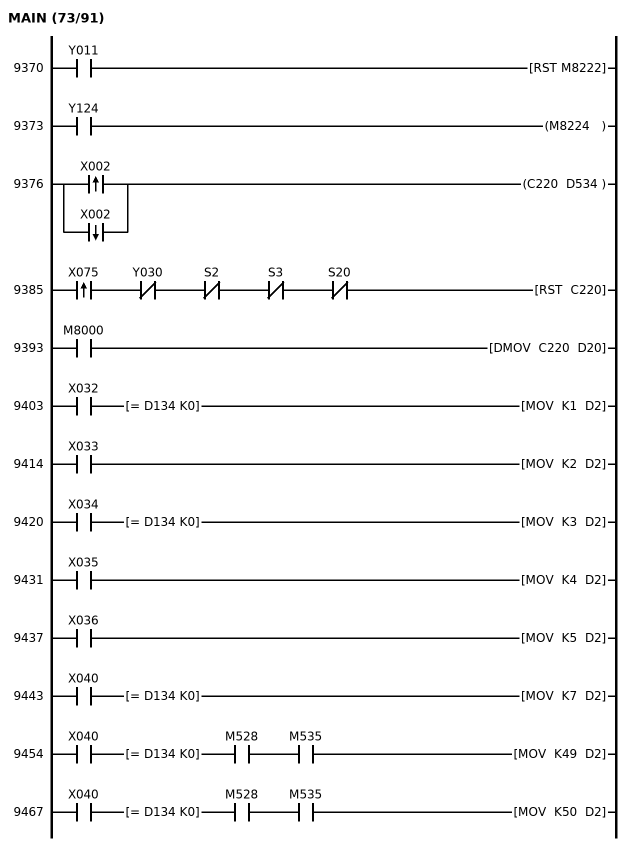
[picture p72: ladder of MAIN, rungs at steps 9370 to 9467]
9370  LD      Y011
      RST     M8222
9373  LD      Y124
      OUT     M8224
9376  LDP     X002
      ORF     X002
      OUT     C220 D534
9385  LDP     X075
      ANI     Y030
      ANI     S2
      ANI     S3
      ANI     S20
      RST     C220
9393  LD      M8000
      DMOV    C220 D20
9403  LD      X032
      AND=    D134 K0
      MOV     K1 D2
9414  LD      X033
      MOV     K2 D2
9420  LD      X034
      AND=    D134 K0
      MOV     K3 D2
9431  LD      X035
      MOV     K4 D2
9437  LD      X036
      MOV     K5 D2
9443  LD      X040
      AND=    D134 K0
      MOV     K7 D2
9454  LD      X040
      AND=    D134 K0
      AND     M528
      AND     M535
      MOV     K49 D2
9467  LD      X040
      AND=    D134 K0
      AND     M528
      AND     M535
      MOV     K50 D2
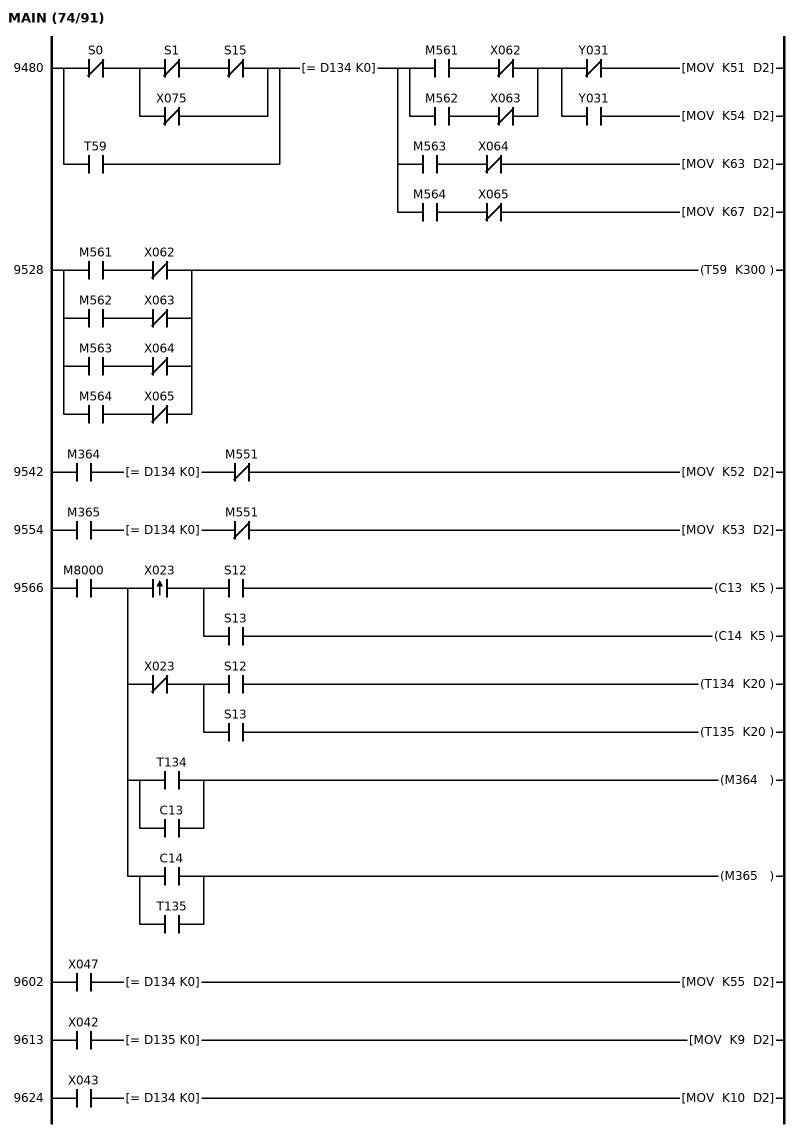
9480  LDI     S0
      LDI     S1
      ANI     S15
      ORI     X075
      ANB
      OR      T59
      AND=    D134 K0
      MPS
      LD      M561
      ANI     X062
      LD      M562
      ANI     X063
      ORB
      ANB
      MPS
      ANI     Y031
      MOV     K51 D2
      MPP
      AND     Y031
      MOV     K54 D2
      MRD
      AND     M563
      ANI     X064
      MOV     K63 D2
      MPP
      AND     M564
      ANI     X065
      MOV     K67 D2
9528  LD      M561
      ANI     X062
      LD      M562
      ANI     X063
      ORB
      LD      M563
      ANI     X064
      ORB
      LD      M564
      ANI     X065
      ORB
      OUT     T59 K300
9542  LD      M364
      AND=    D134 K0
      ANI     M551
      MOV     K52 D2
9554  LD      M365
      AND=    D134 K0
      ANI     M551
      MOV     K53 D2
9566  LD      M8000
      MPS
      ANDP    X023
      MPS
      AND     S12
      OUT     C13 K5
      MPP
      AND     S13
      OUT     C14 K5
      MRD
      ANI     X023
      MPS
      AND     S12
      OUT     T134 K20
      MPP
      AND     S13
      OUT     T135 K20
      MRD
      LD      T134
      OR      C13
      ANB
      OUT     M364
      MPP
      LD      C14
      OR      T135
      ANB
      OUT     M365
9602  LD      X047
      AND=    D134 K0
      MOV     K55 D2
9613  LD      X042
      AND=    D135 K0
      MOV     K9 D2
9624  LD      X043
      AND=    D134 K0
      MOV     K10 D2
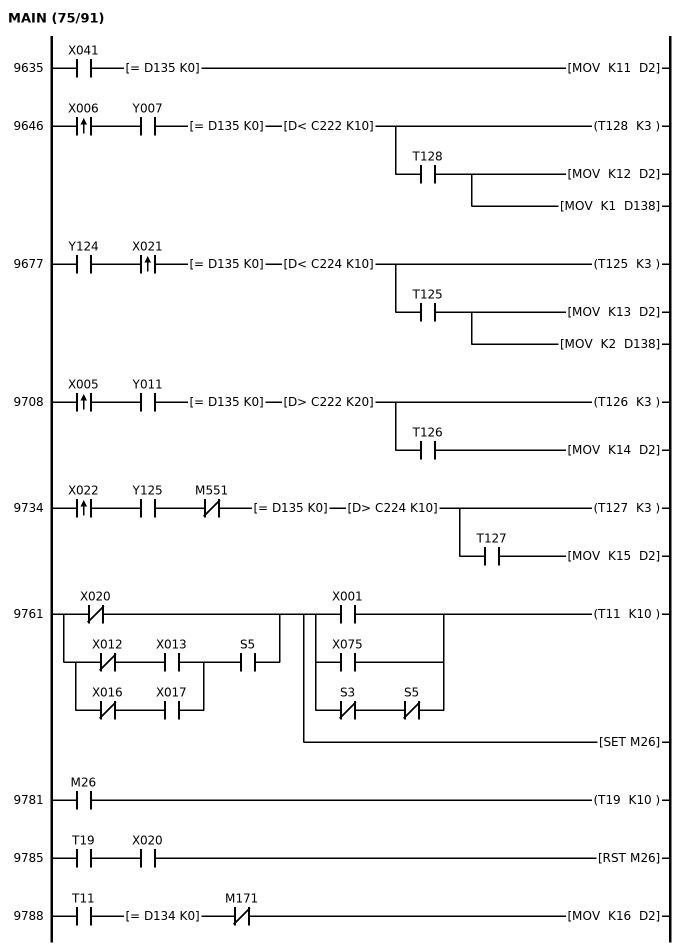
9635  LD      X041
      AND=    D135 K0
      MOV     K11 D2
9646  LDP     X006
      AND     Y007
      AND=    D135 K0
      ANDD<   C222 K10
      OUT     T128 K3
      AND     T128
      MOV     K12 D2
      MOV     K1 D138
9677  LD      Y124
      ANDP    X021
      AND=    D135 K0
      ANDD<   C224 K10
      OUT     T125 K3
      AND     T125
      MOV     K13 D2
      MOV     K2 D138
9708  LDP     X005
      AND     Y011
      AND=    D135 K0
      ANDD>   C222 K20
      OUT     T126 K3
      AND     T126
      MOV     K14 D2
9734  LDP     X022
      AND     Y125
      ANI     M551
      AND=    D135 K0
      ANDD>   C224 K10
      OUT     T127 K3
      AND     T127
      MOV     K15 D2
9761  LDI     X020
      LDI     X012
      AND     X013
      LDI     X016
      AND     X017
      ORB
      AND     S5
      ORB
      MPS
      LD      X001
      OR      X075
      LDI     S3
      ANI     S5
      ORB
      ANB
      OUT     T11 K10
      MPP
      SET     M26
9781  LD      M26
      OUT     T19 K10
9785  LD      T19
      AND     X020
      RST     M26
9788  LD      T11
      AND=    D134 K0
      ANI     M171
      MOV     K16 D2
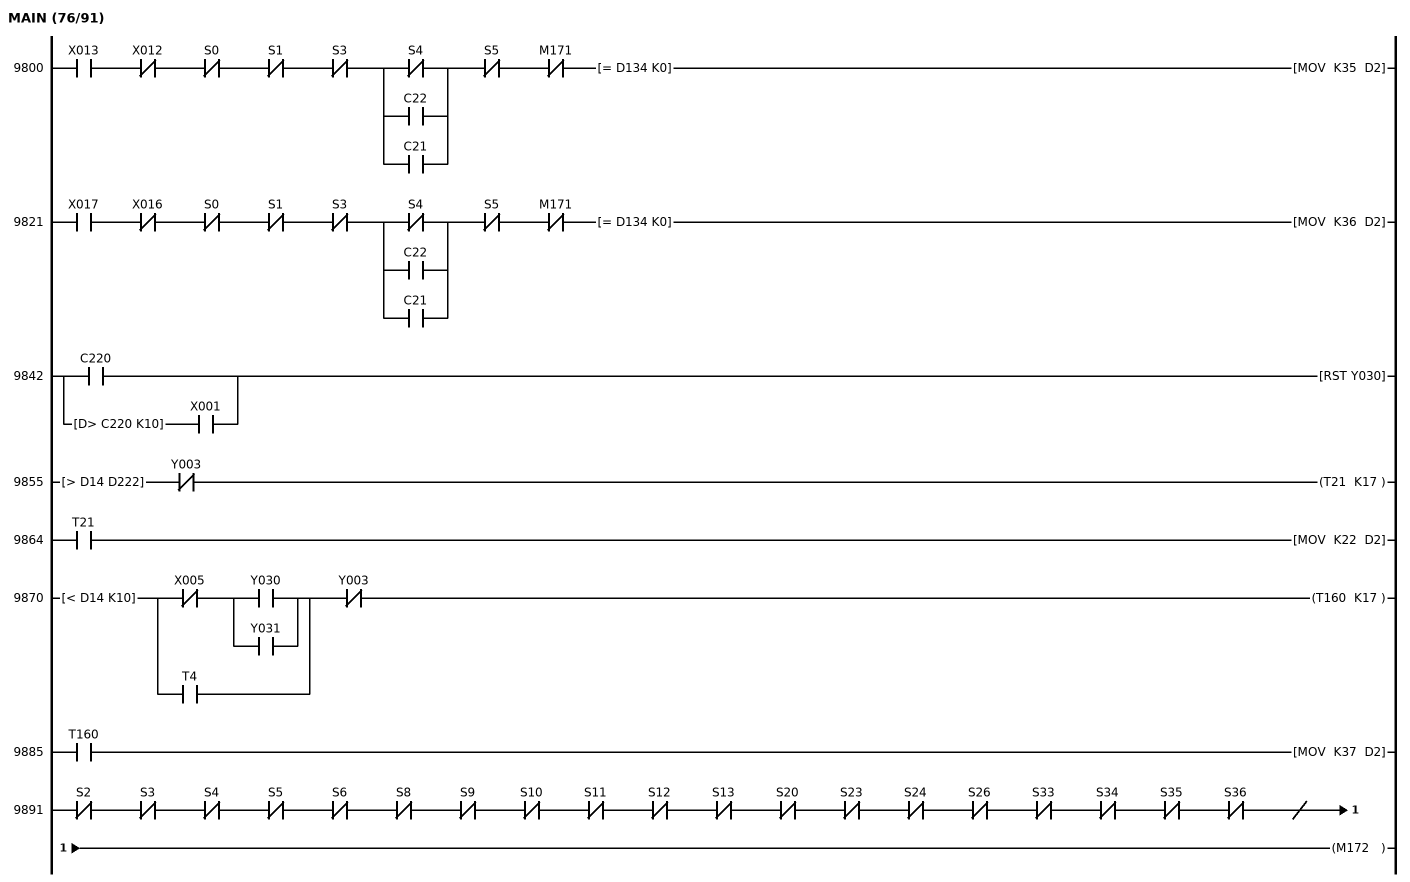
9800  LD      X013
      ANI     X012
      ANI     S0
      ANI     S1
      ANI     S3
      LDI     S4
      OR      C22
      OR      C21
      ANB
      ANI     S5
      ANI     M171
      AND=    D134 K0
      MOV     K35 D2
9821  LD      X017
      ANI     X016
      ANI     S0
      ANI     S1
      ANI     S3
      LDI     S4
      OR      C22
      OR      C21
      ANB
      ANI     S5
      ANI     M171
      AND=    D134 K0
      MOV     K36 D2
9842  LD      C220
      LDD>    C220 K10
      AND     X001
      ORB
      RST     Y030
9855  LD>     D14 D222
      ANI     Y003
      OUT     T21 K17
9864  LD      T21
      MOV     K22 D2
9870  LD<     D14 K10
      LDI     X005
      LD      Y030
      OR      Y031
      ANB
      OR      T4
      ANB
      ANI     Y003
      OUT     T160 K17
9885  LD      T160
      MOV     K37 D2
9891  LDI     S2
      ANI     S3
      ANI     S4
      ANI     S5
      ANI     S6
      ANI     S8
      ANI     S9
      ANI     S10
      ANI     S11
      ANI     S12
      ANI     S13
      ANI     S20
      ANI     S23
      ANI     S24
      ANI     S26
      ANI     S33
      ANI     S34
      ANI     S35
      ANI     S36
      INV
      OUT     M172
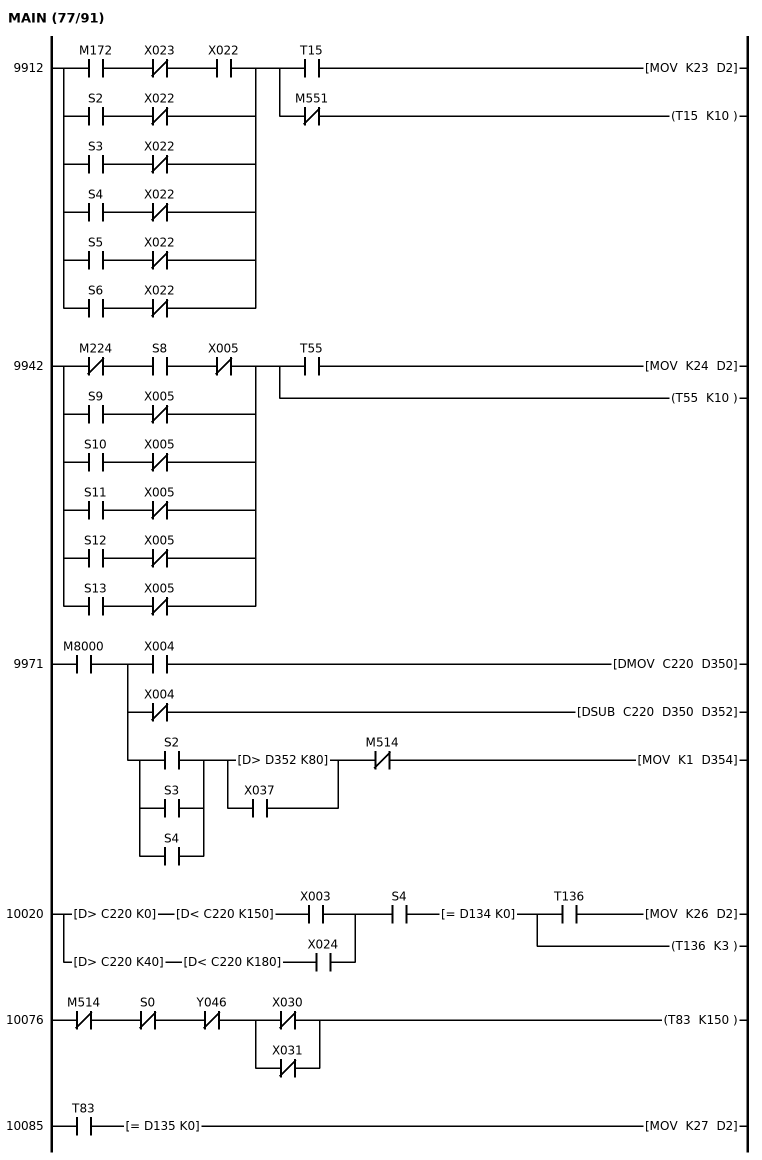
9912  LD      M172
      ANI     X023
      AND     X022
      LD      S2
      ANI     X022
      ORB
      LD      S3
      ANI     X022
      ORB
      LD      S4
      ANI     X022
      ORB
      LD      S5
      ANI     X022
      ORB
      LD      S6
      ANI     X022
      ORB
      MPS
      AND     T15
      MOV     K23 D2
      MPP
      ANI     M551
      OUT     T15 K10
9942  LDI     M224
      AND     S8
      ANI     X005
      LD      S9
      ANI     X005
      ORB
      LD      S10
      ANI     X005
      ORB
      LD      S11
      ANI     X005
      ORB
      LD      S12
      ANI     X005
      ORB
      LD      S13
      ANI     X005
      ORB
      MPS
      AND     T55
      MOV     K24 D2
      MPP
      OUT     T55 K10
9971  LD      M8000
      MPS
      AND     X004
      DMOV    C220 D350
      MRD
      ANI     X004
      DSUB    C220 D350 D352
      MPP
      LD      S2
      OR      S3
      OR      S4
      ANB
      LDD>    D352 K80
      OR      X037
      ANB
      ANI     M514
      MOV     K1 D354
10020 LDD>    C220 K0
      ANDD<   C220 K150
      AND     X003
      LDD>    C220 K40
      ANDD<   C220 K180
      AND     X024
      ORB
      AND     S4
      AND=    D134 K0
      MPS
      AND     T136
      MOV     K26 D2
      MPP
      OUT     T136 K3
10076 LDI     M514
      ANI     S0
      ANI     Y046
      LDI     X030
      ORI     X031
      ANB
      OUT     T83 K150
10085 LD      T83
      AND=    D135 K0
      MOV     K27 D2
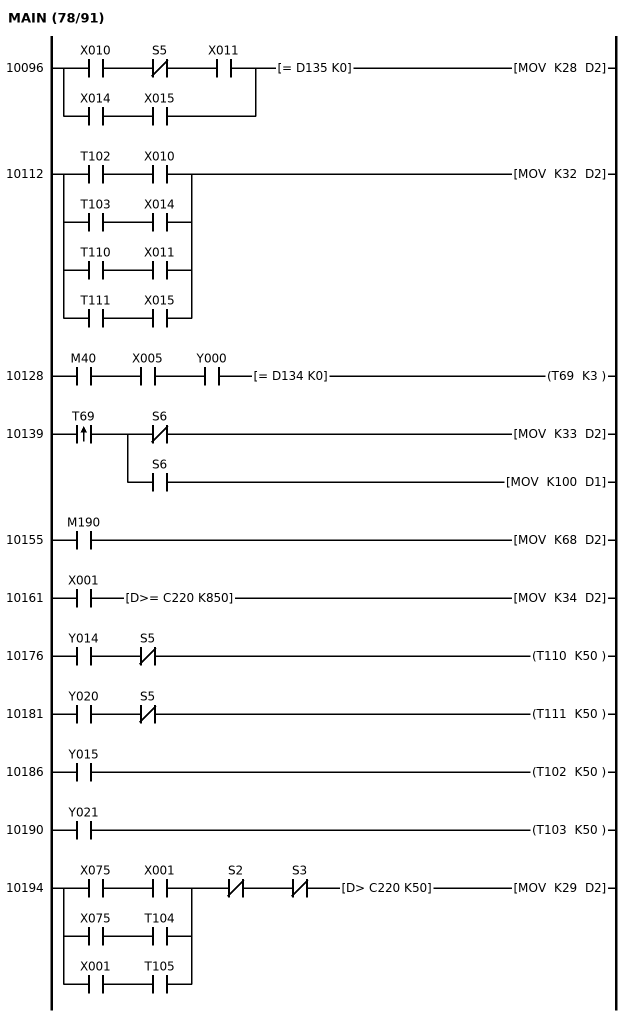
10096 LD      X010
      ANI     S5
      AND     X011
      LD      X014
      AND     X015
      ORB
      AND=    D135 K0
      MOV     K28 D2
10112 LD      T102
      AND     X010
      LD      T103
      AND     X014
      ORB
      LD      T110
      AND     X011
      ORB
      LD      T111
      AND     X015
      ORB
      MOV     K32 D2
10128 LD      M40
      AND     X005
      AND     Y000
      AND=    D134 K0
      OUT     T69 K3
10139 LDP     T69
      MPS
      ANI     S6
      MOV     K33 D2
      MPP
      AND     S6
      MOV     K100 D1
10155 LD      M190
      MOV     K68 D2
10161 LD      X001
      ANDD>=  C220 K850
      MOV     K34 D2
10176 LD      Y014
      ANI     S5
      OUT     T110 K50
10181 LD      Y020
      ANI     S5
      OUT     T111 K50
10186 LD      Y015
      OUT     T102 K50
10190 LD      Y021
      OUT     T103 K50
10194 LD      X075
      AND     X001
      LD      X075
      AND     T104
      ORB
      LD      X001
      AND     T105
      ORB
      ANI     S2
      ANI     S3
      ANDD>   C220 K50
      MOV     K29 D2
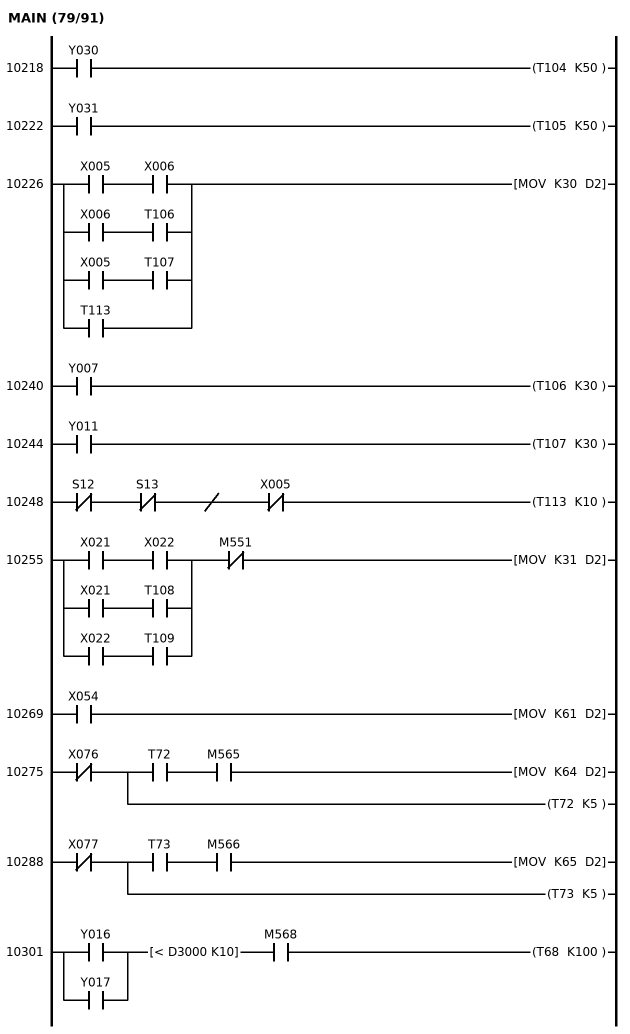
10218 LD      Y030
      OUT     T104 K50
10222 LD      Y031
      OUT     T105 K50
10226 LD      X005
      AND     X006
      LD      X006
      AND     T106
      ORB
      LD      X005
      AND     T107
      ORB
      OR      T113
      MOV     K30 D2
10240 LD      Y007
      OUT     T106 K30
10244 LD      Y011
      OUT     T107 K30
10248 LDI     S12
      ANI     S13
      INV
      ANI     X005
      OUT     T113 K10
10255 LD      X021
      AND     X022
      LD      X021
      AND     T108
      ORB
      LD      X022
      AND     T109
      ORB
      ANI     M551
      MOV     K31 D2
10269 LD      X054
      MOV     K61 D2
10275 LDI     X076
      MPS
      AND     T72
      AND     M565
      MOV     K64 D2
      MPP
      OUT     T72 K5
10288 LDI     X077
      MPS
      AND     T73
      AND     M566
      MOV     K65 D2
      MPP
      OUT     T73 K5
10301 LD      Y016
      OR      Y017
      AND<    D3000 K10
      AND     M568
      OUT     T68 K100
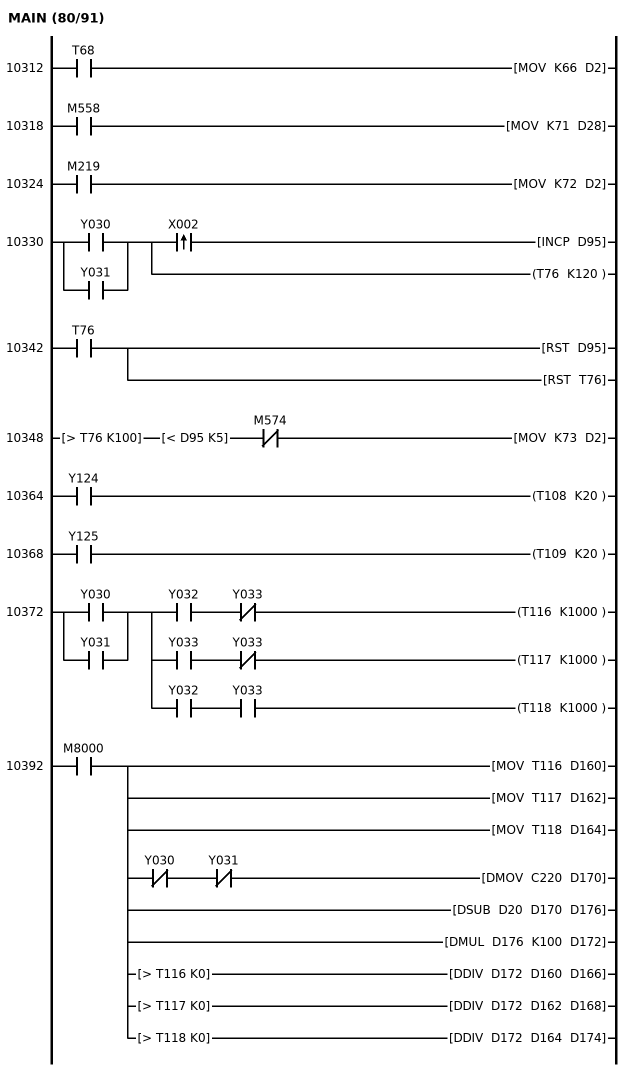
10312 LD      T68
      MOV     K66 D2
10318 LD      M558
      MOV     K71 D28
10324 LD      M219
      MOV     K72 D2
10330 LD      Y030
      OR      Y031
      MPS
      ANDP    X002
      INCP    D95
      MPP
      OUT     T76 K120
10342 LD      T76
      RST     D95
      RST     T76
10348 LD>     T76 K100
      AND<    D95 K5
      ANI     M574
      MOV     K73 D2
10364 LD      Y124
      OUT     T108 K20
10368 LD      Y125
      OUT     T109 K20
10372 LD      Y030
      OR      Y031
      MPS
      AND     Y032
      ANI     Y033
      OUT     T116 K1000
      MRD
      AND     Y033
      ANI     Y033
      OUT     T117 K1000
      MPP
      AND     Y032
      AND     Y033
      OUT     T118 K1000
10392 LD      M8000
      MOV     T116 D160
      MOV     T117 D162
      MOV     T118 D164
      MPS
      ANI     Y030
      ANI     Y031
      DMOV    C220 D170
      MPP
      DSUB    D20 D170 D176
      DMUL    D176 K100 D172
      MPS
      AND>    T116 K0
      DDIV    D172 D160 D166
      MRD
      AND>    T117 K0
      DDIV    D172 D162 D168
      MPP
      AND>    T118 K0
      DDIV    D172 D164 D174
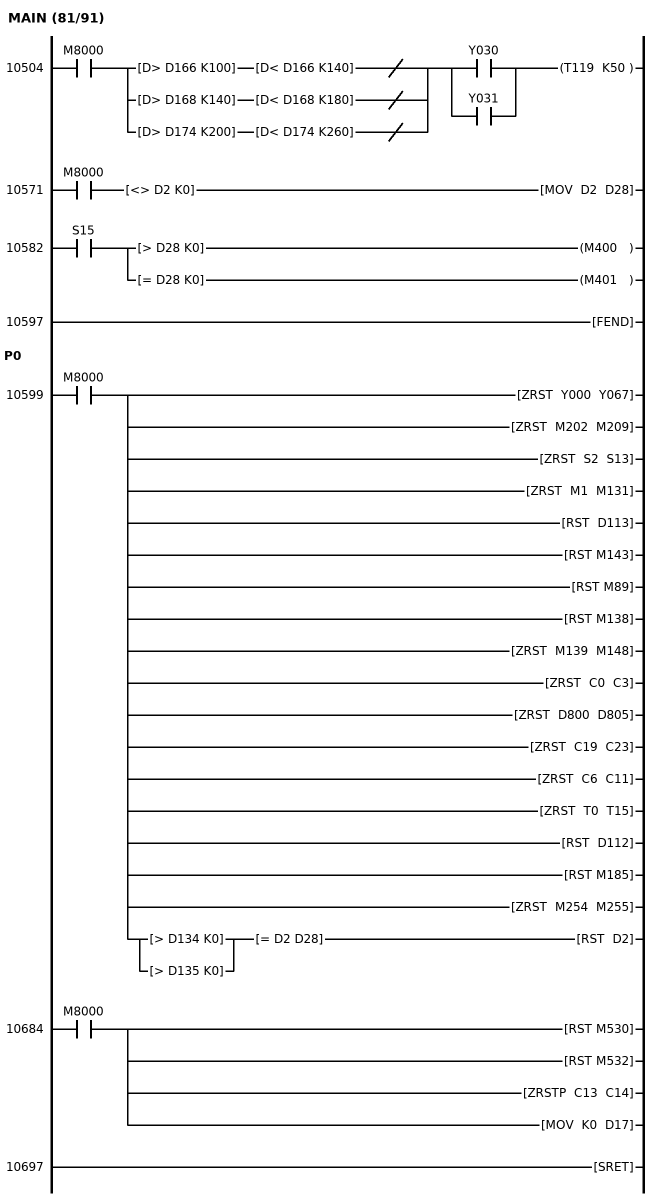
10504 LD      M8000
      LDD>    D166 K100
      ANDD<   D166 K140
      INV
      LDD>    D168 K140
      ANDD<   D168 K180
      INV
      ORB
      LDD>    D174 K200
      ANDD<   D174 K260
      INV
      ORB
      ANB
      LD      Y030
      OR      Y031
      ANB
      OUT     T119 K50
10571 LD      M8000
      AND<>   D2 K0
      MOV     D2 D28
10582 LD      S15
      MPS
      AND>    D28 K0
      OUT     M400
      MPP
      AND=    D28 K0
      OUT     M401
10597 FEND
      P0
10599 LD      M8000
      ZRST    Y000 Y067
      ZRST    M202 M209
      ZRST    S2 S13
      ZRST    M1 M131
      RST     D113
      RST     M143
      RST     M89
      RST     M138
      ZRST    M139 M148
      ZRST    C0 C3
      ZRST    D800 D805
      ZRST    C19 C23
      ZRST    C6 C11
      ZRST    T0 T15
      RST     D112
      RST     M185
      ZRST    M254 M255
      LD>     D134 K0
      OR>     D135 K0
      ANB
      AND=    D2 D28
      RST     D2
10684 LD      M8000
      RST     M530
      RST     M532
      ZRSTP   C13 C14
      MOV     K0 D17
10697 SRET
      P1
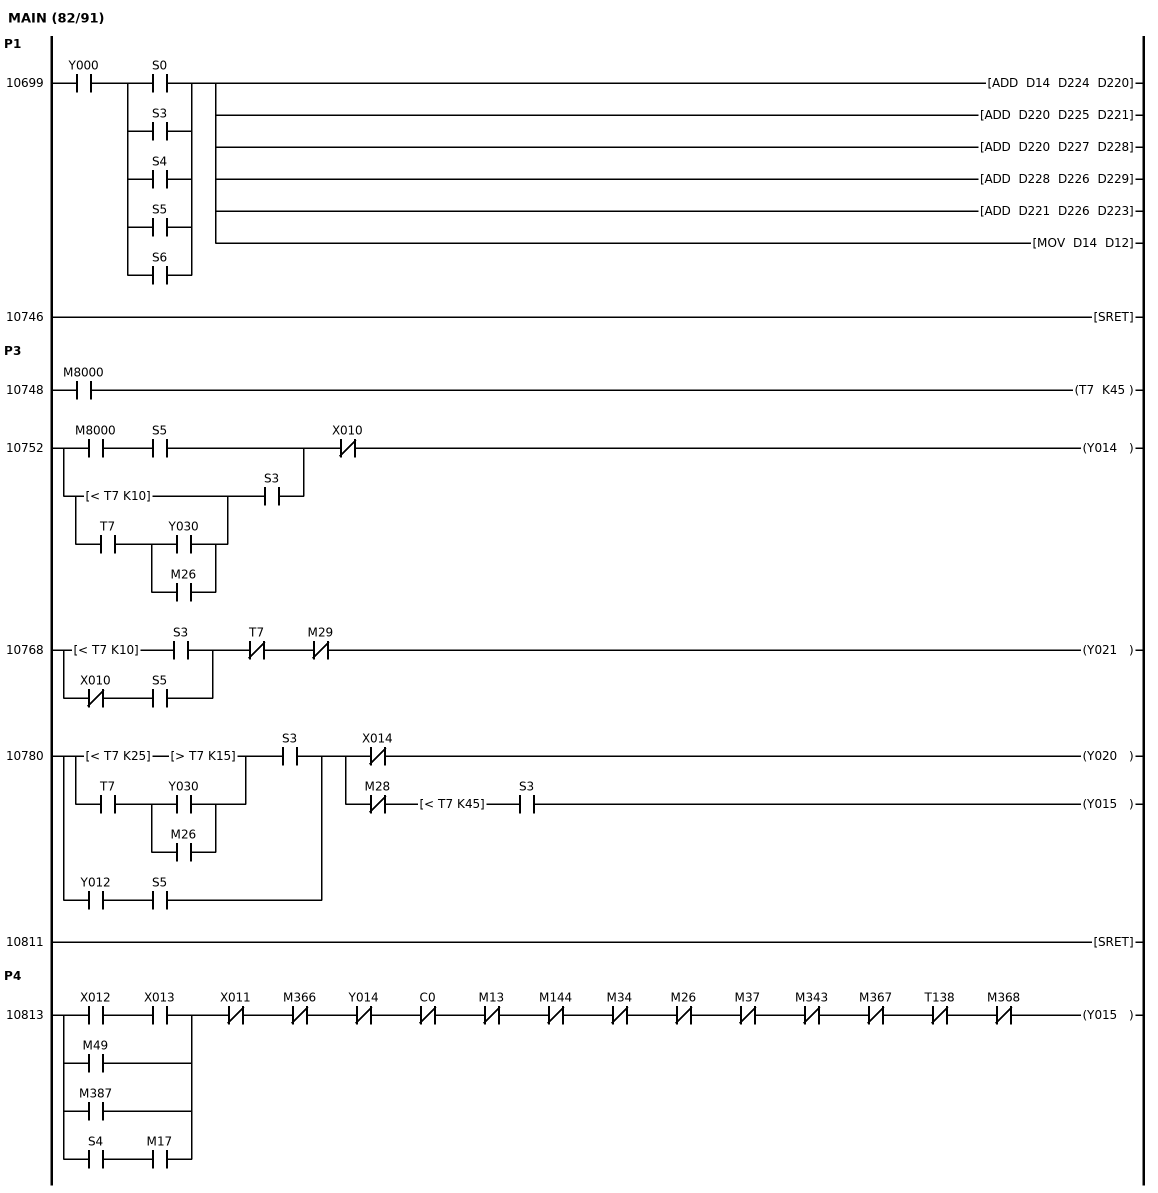
10699 LD      Y000
      LD      S0
      OR      S3
      OR      S4
      OR      S5
      OR      S6
      ANB
      ADD     D14 D224 D220
      ADD     D220 D225 D221
      ADD     D220 D227 D228
      ADD     D228 D226 D229
      ADD     D221 D226 D223
      MOV     D14 D12
10746 SRET
      P3
10748 LD      M8000
      OUT     T7 K45
10752 LD      M8000
      AND     S5
      LD<     T7 K10
      LD      T7
      LD      Y030
      OR      M26
      ANB
      ORB
      AND     S3
      ORB
      ANI     X010
      OUT     Y014
10768 LD<     T7 K10
      AND     S3
      LDI     X010
      AND     S5
      ORB
      ANI     T7
      ANI     M29
      OUT     Y021
10780 LD<     T7 K25
      AND>    T7 K15
      LD      T7
      LD      Y030
      OR      M26
      ANB
      ORB
      AND     S3
      LD      Y012
      AND     S5
      ORB
      MPS
      ANI     X014
      OUT     Y020
      MPP
      ANI     M28
      AND<    T7 K45
      AND     S3
      OUT     Y015
10811 SRET
      P4
10813 LD      X012
      AND     X013
      OR      M49
      OR      M387
      LD      S4
      AND     M17
      ORB
      ANI     X011
      ANI     M366
      ANI     Y014
      ANI     C0
      ANI     M13
      ANI     M144
      ANI     M34
      ANI     M26
      ANI     M37
      ANI     M343
      ANI     M367
      ANI     T138
      ANI     M368
      OUT     Y015
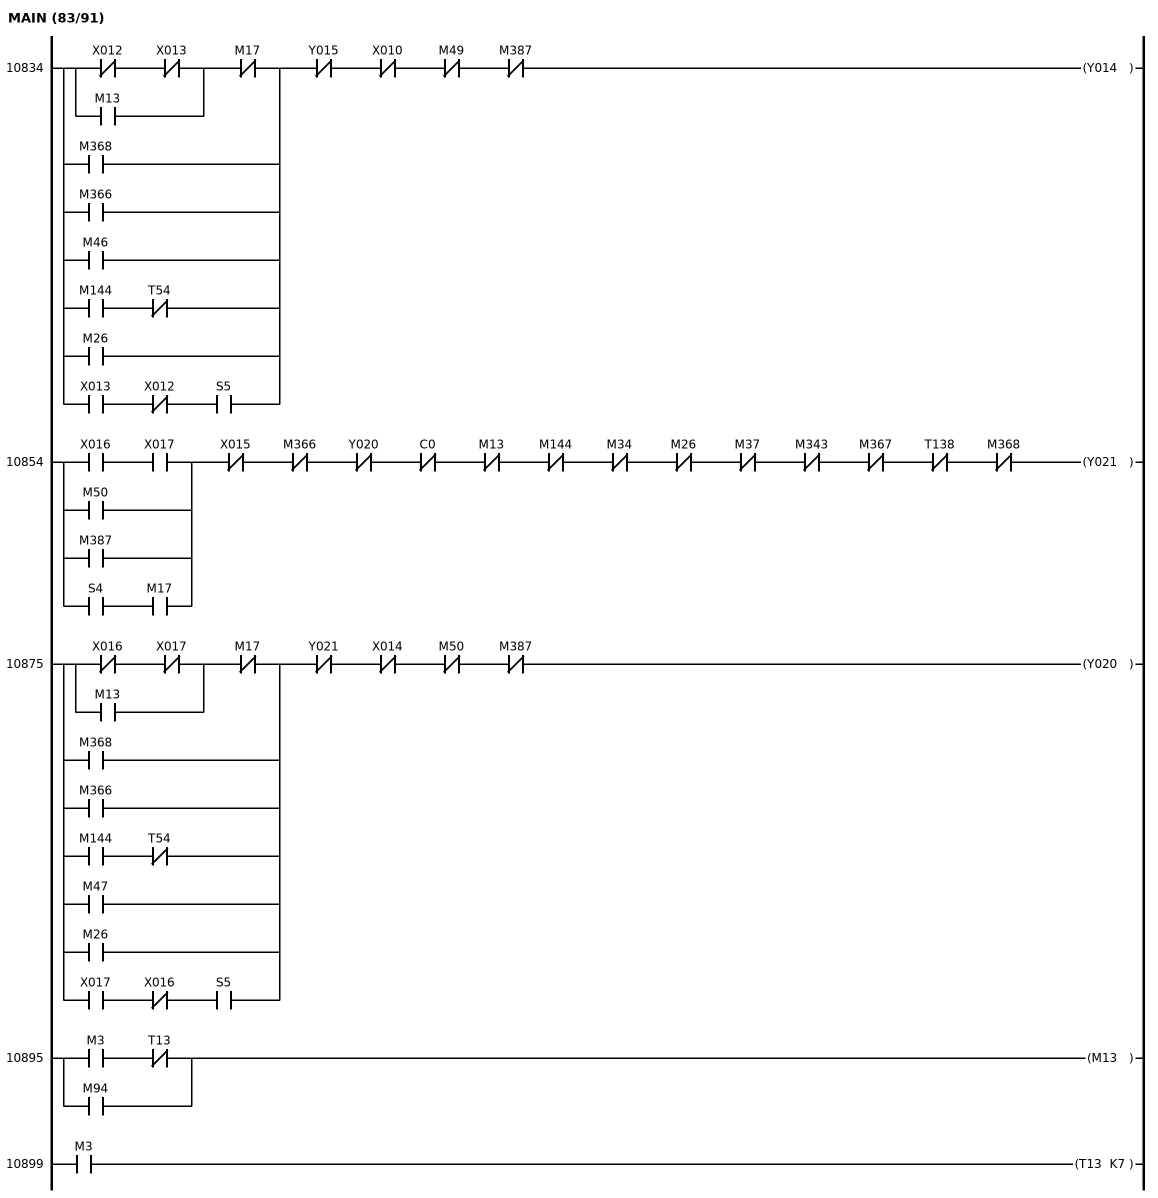
10834 LDI     X012
      ANI     X013
      OR      M13
      ANI     M17
      OR      M368
      OR      M366
      OR      M46
      LD      M144
      ANI     T54
      ORB
      OR      M26
      LD      X013
      ANI     X012
      AND     S5
      ORB
      ANI     Y015
      ANI     X010
      ANI     M49
      ANI     M387
      OUT     Y014
10854 LD      X016
      AND     X017
      OR      M50
      OR      M387
      LD      S4
      AND     M17
      ORB
      ANI     X015
      ANI     M366
      ANI     Y020
      ANI     C0
      ANI     M13
      ANI     M144
      ANI     M34
      ANI     M26
      ANI     M37
      ANI     M343
      ANI     M367
      ANI     T138
      ANI     M368
      OUT     Y021
10875 LDI     X016
      ANI     X017
      OR      M13
      ANI     M17
      OR      M368
      OR      M366
      LD      M144
      ANI     T54
      ORB
      OR      M47
      OR      M26
      LD      X017
      ANI     X016
      AND     S5
      ORB
      ANI     Y021
      ANI     X014
      ANI     M50
      ANI     M387
      OUT     Y020
10895 LD      M3
      ANI     T13
      OR      M94
      OUT     M13
10899 LD      M3
      OUT     T13 K7
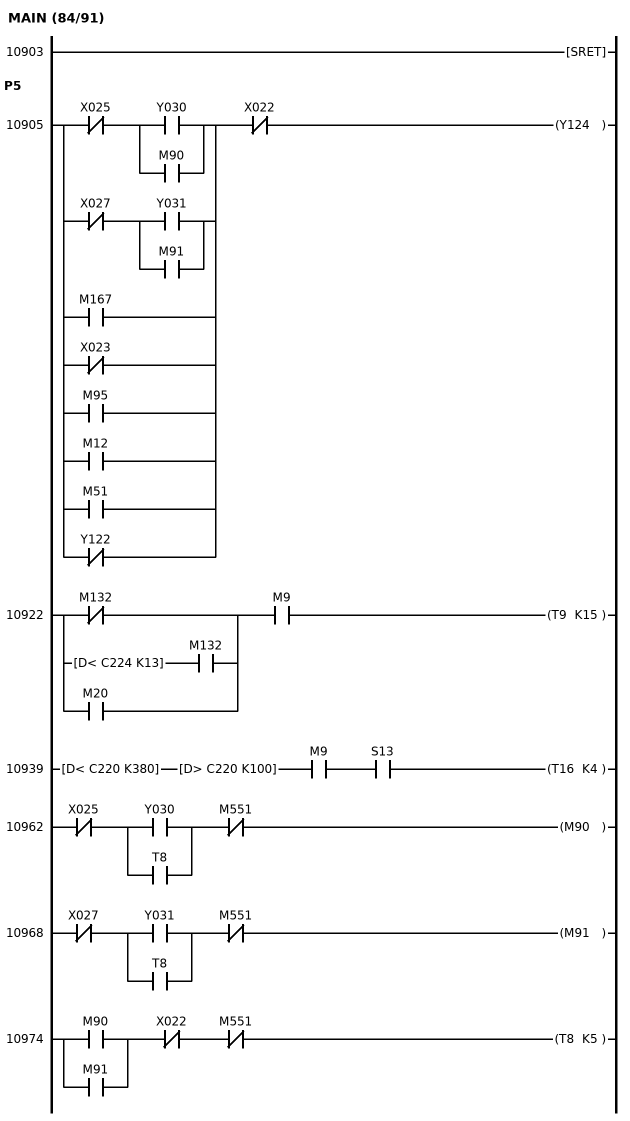
10903 SRET
      P5
10905 LDI     X025
      LD      Y030
      OR      M90
      ANB
      LDI     X027
      LD      Y031
      OR      M91
      ANB
      ORB
      OR      M167
      ORI     X023
      OR      M95
      OR      M12
      OR      M51
      ORI     Y122
      ANI     X022
      OUT     Y124
10922 LDI     M132
      LDD<    C224 K13
      AND     M132
      ORB
      OR      M20
      AND     M9
      OUT     T9 K15
10939 LDD<    C220 K380
      ANDD>   C220 K100
      AND     M9
      AND     S13
      OUT     T16 K4
10962 LDI     X025
      LD      Y030
      OR      T8
      ANB
      ANI     M551
      OUT     M90
10968 LDI     X027
      LD      Y031
      OR      T8
      ANB
      ANI     M551
      OUT     M91
10974 LD      M90
      OR      M91
      ANI     X022
      ANI     M551
      OUT     T8 K5
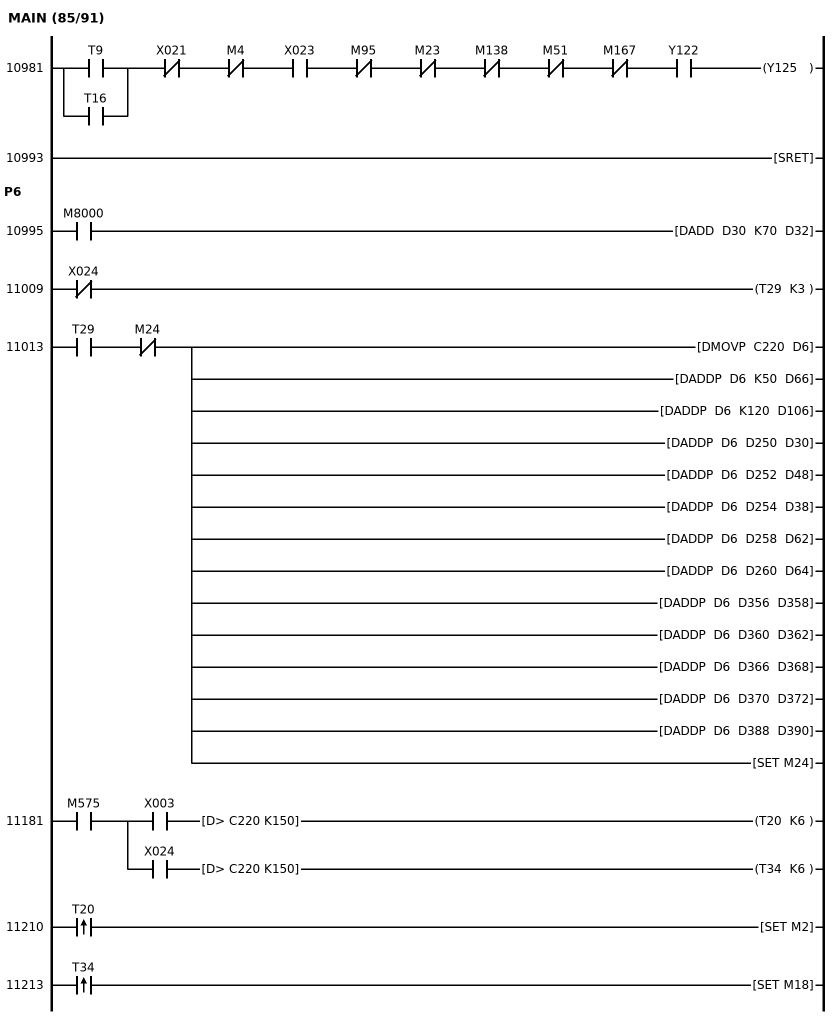
10981 LD      T9
      OR      T16
      ANI     X021
      ANI     M4
      AND     X023
      ANI     M95
      ANI     M23
      ANI     M138
      ANI     M51
      ANI     M167
      AND     Y122
      OUT     Y125
10993 SRET
      P6
10995 LD      M8000
      DADD    D30 K70 D32
11009 LDI     X024
      OUT     T29 K3
11013 LD      T29
      ANI     M24
      DMOVP   C220 D6
      DADDP   D6 K50 D66
      DADDP   D6 K120 D106
      DADDP   D6 D250 D30
      DADDP   D6 D252 D48
      DADDP   D6 D254 D38
      DADDP   D6 D258 D62
      DADDP   D6 D260 D64
      DADDP   D6 D356 D358
      DADDP   D6 D360 D362
      DADDP   D6 D366 D368
      DADDP   D6 D370 D372
      DADDP   D6 D388 D390
      SET     M24
11181 LD      M575
      MPS
      AND     X003
      ANDD>   C220 K150
      OUT     T20 K6
      MPP
      AND     X024
      ANDD>   C220 K150
      OUT     T34 K6
11210 LDP     T20
      SET     M2
11213 LDP     T34
      SET     M18
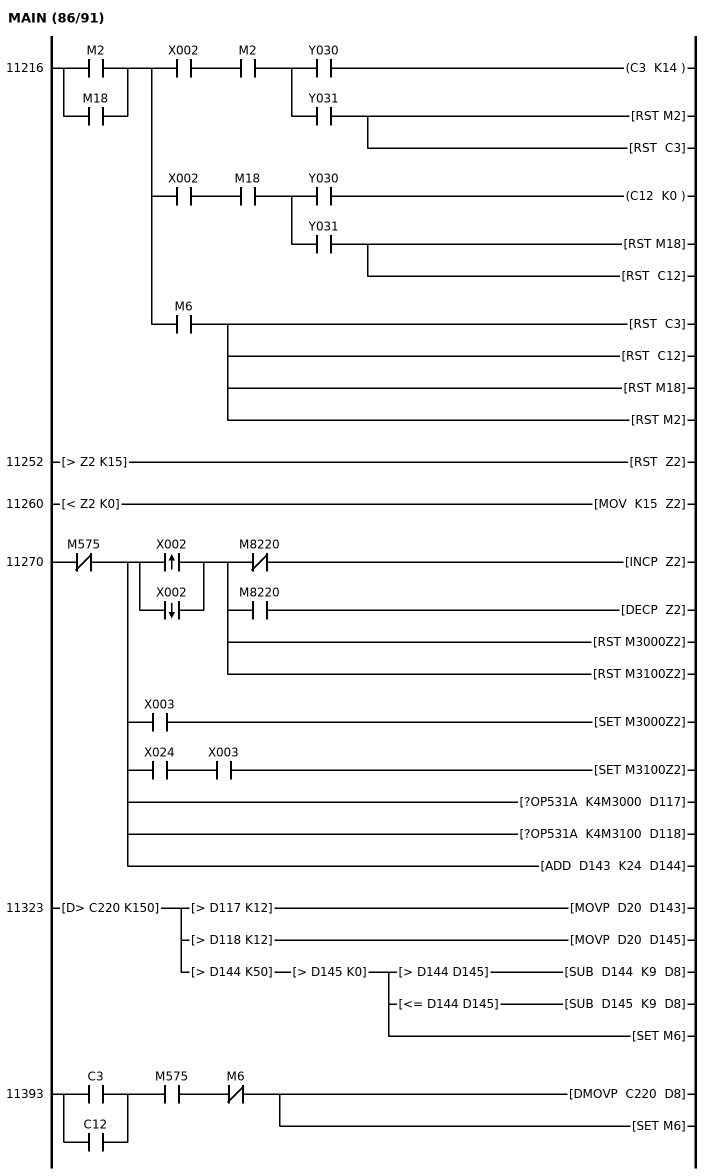
11216 LD      M2
      OR      M18
      MPS
      AND     X002
      AND     M2
      MPS
      AND     Y030
      OUT     C3 K14
      MPP
      AND     Y031
      RST     M2
      RST     C3
      MRD
      AND     X002
      AND     M18
      MPS
      AND     Y030
      OUT     C12 K0
      MPP
      AND     Y031
      RST     M18
      RST     C12
      MPP
      AND     M6
      RST     C3
      RST     C12
      RST     M18
      RST     M2
11252 LD>     Z2 K15
      RST     Z2
11260 LD<     Z2 K0
      MOV     K15 Z2
11270 LDI     M575
      MPS
      LDP     X002
      ORF     X002
      ANB
      MPS
      ANI     M8220
      INCP    Z2
      MRD
      AND     M8220
      DECP    Z2
      MPP
      RST     M3000Z2
      RST     M3100Z2
      MRD
      AND     X003
      SET     M3000Z2
      MRD
      AND     X024
      AND     X003
      SET     M3100Z2
      MPP
      ?OP531A K4M3000 D117
      ?OP531A K4M3100 D118
      ADD     D143 K24 D144
11323 LDD>    C220 K150
      MPS
      AND>    D117 K12
      MOVP    D20 D143
      MRD
      AND>    D118 K12
      MOVP    D20 D145
      MPP
      AND>    D144 K50
      AND>    D145 K0
      MPS
      AND>    D144 D145
      SUB     D144 K9 D8
      MRD
      AND<=   D144 D145
      SUB     D145 K9 D8
      MPP
      SET     M6
11393 LD      C3
      OR      C12
      AND     M575
      ANI     M6
      DMOVP   C220 D8
      SET     M6
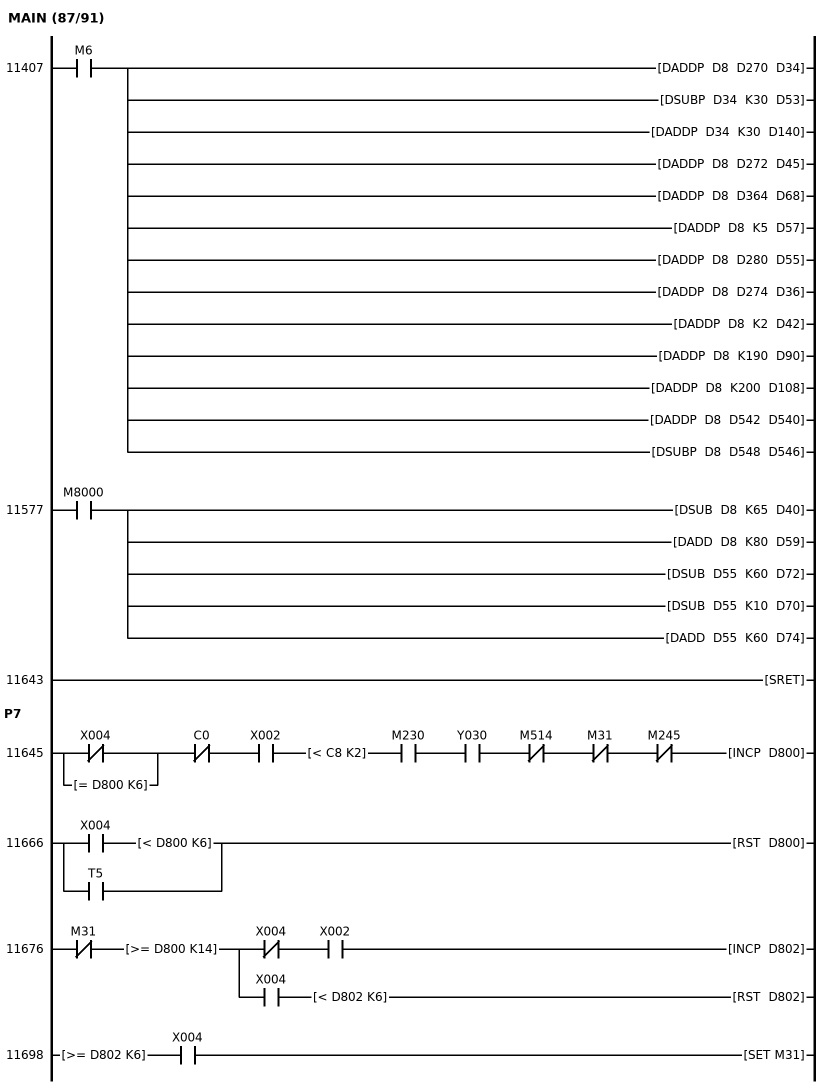
11407 LD      M6
      DADDP   D8 D270 D34
      DSUBP   D34 K30 D53
      DADDP   D34 K30 D140
      DADDP   D8 D272 D45
      DADDP   D8 D364 D68
      DADDP   D8 K5 D57
      DADDP   D8 D280 D55
      DADDP   D8 D274 D36
      DADDP   D8 K2 D42
      DADDP   D8 K190 D90
      DADDP   D8 K200 D108
      DADDP   D8 D542 D540
      DSUBP   D8 D548 D546
11577 LD      M8000
      DSUB    D8 K65 D40
      DADD    D8 K80 D59
      DSUB    D55 K60 D72
      DSUB    D55 K10 D70
      DADD    D55 K60 D74
11643 SRET
      P7
11645 LDI     X004
      OR=     D800 K6
      ANI     C0
      AND     X002
      AND<    C8 K2
      AND     M230
      AND     Y030
      ANI     M514
      ANI     M31
      ANI     M245
      INCP    D800
11666 LD      X004
      AND<    D800 K6
      OR      T5
      RST     D800
11676 LDI     M31
      AND>=   D800 K14
      MPS
      ANI     X004
      AND     X002
      INCP    D802
      MPP
      AND     X004
      AND<    D802 K6
      RST     D802
11698 LD>=    D802 K6
      AND     X004
      SET     M31
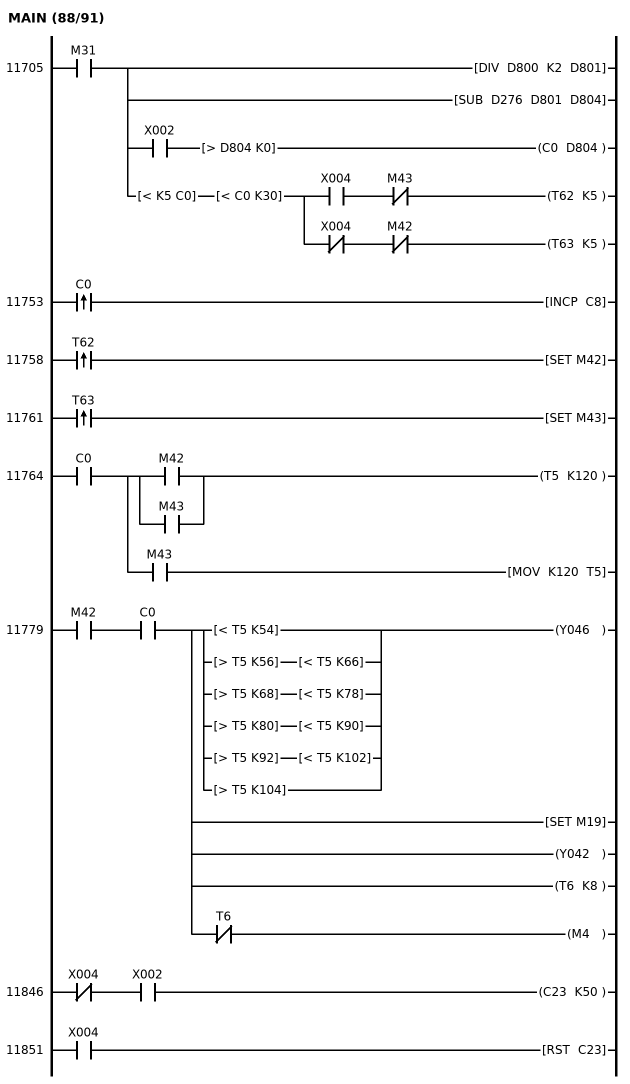
11705 LD      M31
      DIV     D800 K2 D801
      SUB     D276 D801 D804
      MPS
      AND     X002
      AND>    D804 K0
      OUT     C0 D804
      MPP
      AND<    K5 C0
      AND<    C0 K30
      MPS
      AND     X004
      ANI     M43
      OUT     T62 K5
      MPP
      ANI     X004
      ANI     M42
      OUT     T63 K5
11753 LDP     C0
      INCP    C8
11758 LDP     T62
      SET     M42
11761 LDP     T63
      SET     M43
11764 LD      C0
      MPS
      LD      M42
      OR      M43
      ANB
      OUT     T5 K120
      MPP
      AND     M43
      MOV     K120 T5
11779 LD      M42
      AND     C0
      MPS
      LD<     T5 K54
      LD>     T5 K56
      AND<    T5 K66
      ORB
      LD>     T5 K68
      AND<    T5 K78
      ORB
      LD>     T5 K80
      AND<    T5 K90
      ORB
      LD>     T5 K92
      AND<    T5 K102
      ORB
      OR>     T5 K104
      ANB
      OUT     Y046
      MPP
      SET     M19
      OUT     Y042
      OUT     T6 K8
      ANI     T6
      OUT     M4
11846 LDI     X004
      AND     X002
      OUT     C23 K50
11851 LD      X004
      RST     C23
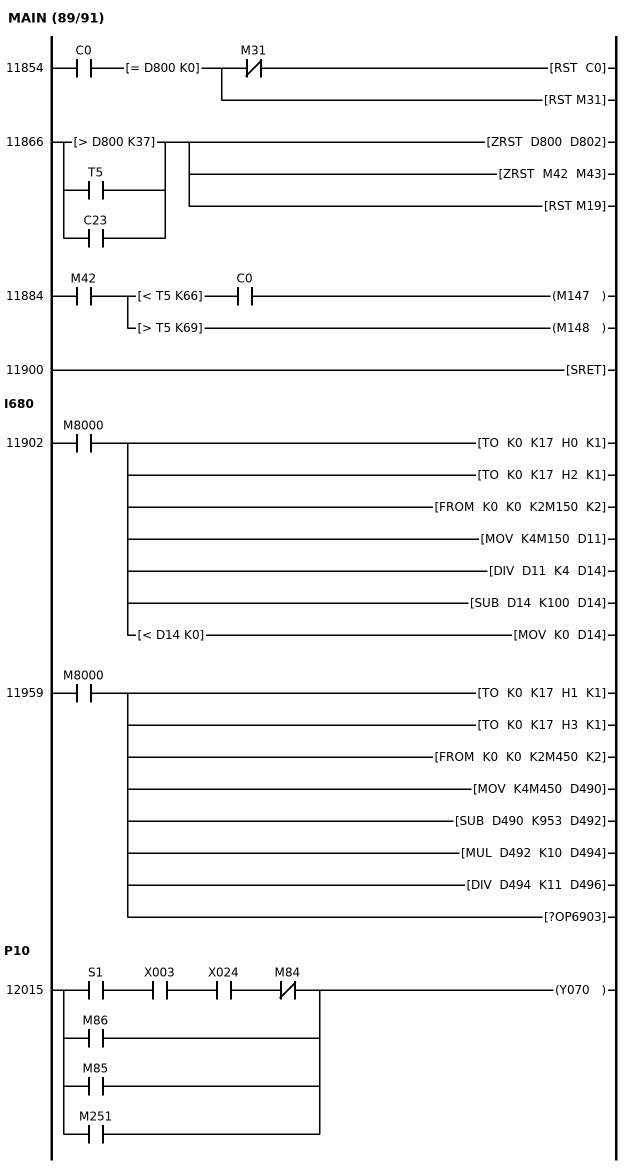
11854 LD      C0
      AND=    D800 K0
      MPS
      ANI     M31
      RST     C0
      MPP
      RST     M31
11866 LD>     D800 K37
      OR      T5
      OR      C23
      ZRST    D800 D802
      ZRST    M42 M43
      RST     M19
11884 LD      M42
      MPS
      AND<    T5 K66
      AND     C0
      OUT     M147
      MPP
      AND>    T5 K69
      OUT     M148
11900 SRET
      I680
11902 LD      M8000
      TO      K0 K17 H0 K1
      TO      K0 K17 H2 K1
      FROM    K0 K0 K2M150 K2
      MOV     K4M150 D11
      DIV     D11 K4 D14
      SUB     D14 K100 D14
      AND<    D14 K0
      MOV     K0 D14
11959 LD      M8000
      TO      K0 K17 H1 K1
      TO      K0 K17 H3 K1
      FROM    K0 K0 K2M450 K2
      MOV     K4M450 D490
      SUB     D490 K953 D492
      MUL     D492 K10 D494
      DIV     D494 K11 D496
      ?OP6903
      P10
12015 LD      S1
      AND     X003
      AND     X024
      ANI     M84
      OR      M86
      OR      M85
      OR      M251
      OUT     Y070
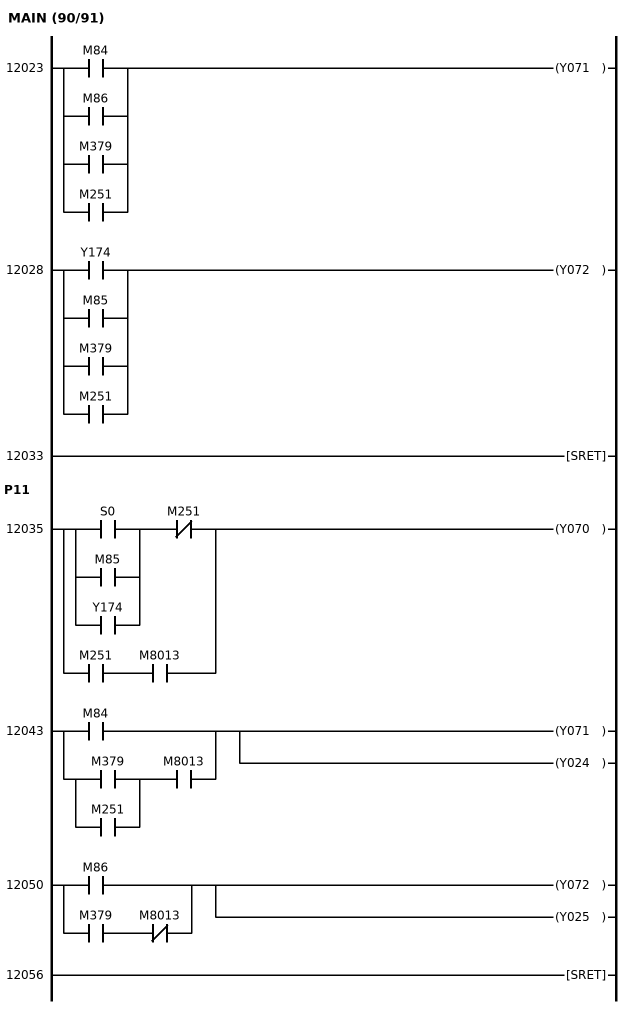
12023 LD      M84
      OR      M86
      OR      M379
      OR      M251
      OUT     Y071
12028 LD      Y174
      OR      M85
      OR      M379
      OR      M251
      OUT     Y072
12033 SRET
      P11
12035 LD      S0
      OR      M85
      OR      Y174
      ANI     M251
      LD      M251
      AND     M8013
      ORB
      OUT     Y070
12043 LD      M84
      LD      M379
      OR      M251
      AND     M8013
      ORB
      OUT     Y071
      OUT     Y024
12050 LD      M86
      LD      M379
      ANI     M8013
      ORB
      OUT     Y072
      OUT     Y025
12056 SRET
      P12
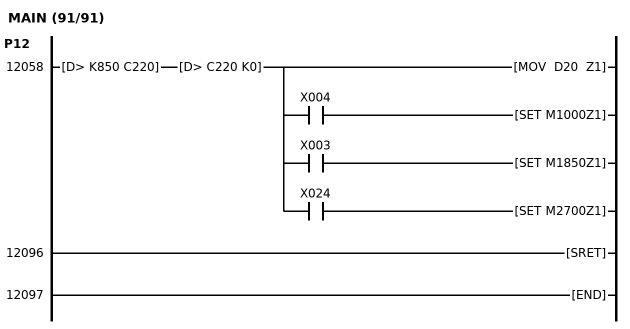
12058 LDD>    K850 C220
      ANDD>   C220 K0
      MOV     D20 Z1
      MPS
      AND     X004
      SET     M1000Z1
      MRD
      AND     X003
      SET     M1850Z1
      MPP
      AND     X024
      SET     M2700Z1
12096 SRET
12097 END
END_PROGRAM
